// TIA Portal V21 export
// export: Created 2026-10-14T03:08:59.3393897Z, ExportSetting WithDefaults, DisplayName Totally Integrated Automation Portal, DisplayVersion V21, DisplayName STEP 7 Professional, DisplayVersion V21, DisplayName STEP 7 Safety, DisplayVersion V21, DisplayName Tech WebApplication, DisplayVersion V21, DisplayName WinCC Basic/Comfort/Advanced, DisplayVersion V21, DisplayName WinCC Unified, DisplayVersion V21
VAR_GLOBAL   // PLC tag table "Default tag table"
   Manipulator AT %MW0 : Int;
END_VAR
VAR_GLOBAL CONSTANT   // user constants
   STATE_FILL_TANK : Int := 1;
   STATE_HEAT_TANK : Int := 2;
   STATE_FILL_BOTTLE : Int := 3;
   STATE_SHIFT_BOTTLE : Int := 4;
   STATE_STOP : Int := 5;
   STATE_RESET : Int := 6;
   STATE_ERROR : Int := 7;
   ERROR_0_NoError : UInt := 8000;
   ERROR_1_BottleInWrongPosition : UInt := 8001;
   ERROR_2_CrackedBottleDetected : UInt := 8002;
   ERROR_3_NoBottleOnTheConveyor : UInt := 8003;
   ERROR_4_WrongBottleDetected : UInt := 8004;
   ERROR_5_ConveyorMalfunction : UInt := 8005;
   ERROR_6_FillerMalfunction : UInt := 8006;
   ERROR_7_ValveBlocked : UInt := 8007;
   ERROR_8_NoFlowInMainPipe : UInt := 8008;
   ERROR_9_GenericError_CheckPlcBuffer : UInt := 8009;
   ERROR_10_GenericError_CheckAlarmBuffer : UInt := 8010;
   ERROR_11_GenericError_ContactWithSupplier : UInt := 8011;
   OEE_ERROR_1_BottleInWrongPosition : UInt := 4;
   OEE_ERROR_10_GenericError_CheckAlarmBuffer : UInt := 13;
   OEE_ERROR_11_GenericError_ContactWithSupplier : UInt := 14;
   OEE_ERROR_2_CrackedBottleDetected : UInt := 5;
   OEE_ERROR_3_NoBottleOnTheConveyor : UInt := 6;
   OEE_ERROR_4_WrongBottleDetected : UInt := 7;
   OEE_ERROR_5_ConveyorMalfunction : UInt := 8;
   OEE_ERROR_6_FillerMalfunction : UInt := 9;
   OEE_ERROR_7_ValveBlocked : UInt := 10;
   OEE_ERROR_8_NoFlowInMainPipe : UInt := 11;
   OEE_ERROR_9_GenericError_CheckPlcBuffer : UInt := 12;
   OEE_PRODUCTION : UInt := 1;
   OEE_PLANNED_DOWN : UInt := 2;
   OEE_UNPLANNED_DOWN : UInt := 3;
END_VAR
